FUNCTION_BLOCK TcoObjectTest EXTENDS TcoCore.TcoObject
VAR
	_myIdentity				:	ULINT;
	_myContextIdentity		:	ULINT;
	_myContextStartCount 	:	ULINT;
	_myContextEndCount		:	ULINT;
	_myParentIdentity		:	ULINT;
	_tcoTaskTest_A			:	TcoTaskTest(THIS^);
	_tcoTaskTest_B			:	TcoTaskTest(THIS^);
	_tcoStateTest_A			:	TcoStateTest(THIS^, eRestoreMode.AutoRestoreMembers);
	_tcoStateTest_B			:	TcoStateTest(THIS^, eRestoreMode.None);
	// Object equality
	_tcoObjectEqualsTestObj1 	:   TcoObjectEqualsTest(THIS^);
	_tcoObjectEqualsTestObj2 	:   TcoObjectEqualsTest(THIS^);
END_VAR

{attribute 'TcRpcEnable'}
METHOD INTERNAL CallTaskInstancies
_tcoTaskTest_A();

_tcoTaskTest_B();
END_METHOD

{attribute 'TcRpcEnable'}
METHOD PUBLIC EqualsOverrideTest : BOOL
EqualsOverrideTest := _tcoObjectEqualsTestObj1.EqualsTo(_tcoObjectEqualsTestObj2);
END_METHOD

{attribute 'TcRpcEnable'}
METHOD PUBLIC EqualsTest : BOOL
VAR_INPUT
    _case : INT;
END_VAR

VAR
    referenceTo_a_TcoStateTest : REFERENCE TO TcoStateTest;
END_VAR
CASE _case OF
    0:
        referenceTo_a_TcoStateTest REF= _tcoStateTest_A;
        EqualsTest := _tcoStateTest_A.EqualsTo(referenceTo_a_TcoStateTest);
    1:
        EqualsTest := _tcoStateTest_A.EqualsTo(_tcoStateTest_B);
    4:
        EqualsTest := _tcoStateTest_B.EqualsTo(_tcoStateTest_A);
    2:
        EqualsTest := _tcoObjectEqualsTestObj1.EqualsTo(_tcoObjectEqualsTestObj1);
    3:
        EqualsTest := _tcoObjectEqualsTestObj1.EqualsTo(_tcoObjectEqualsTestObj2);
END_CASE
END_METHOD

{attribute 'TcRpcEnable'}
METHOD INTERNAL ReadOutIdentities
_myIdentity			:=	THIS^.Identity;

_myContextIdentity	:=	THIS^.Context.Identity;
		
_myContextStartCount :=	THIS^.Context.StartCycleCount;

_myContextEndCount	:=	THIS^.Context.EndCycleCount;

_myParentIdentity	:=	THIS^.Parent.Identity;
END_METHOD

END_FUNCTION_BLOCK

(* stored: Version 1.1.0.1
   POU TcoObjectTest: Id {e84228ff-9c33-47a4-a38e-640688a82a88}, SpecialFunc None
   Method CallTaskInstancies: Id {ca9ba4d2-6103-4337-95bc-465f8f83317e}
   Method EqualsOverrideTest: Id {ee60d2fd-b5db-0d20-0c27-57a751cde2ce}
   Method EqualsTest: Id {9f06ff61-1678-0fe4-0121-54cfb8b16218}
   Method ReadOutIdentities: Id {b42bfa48-43e7-40ad-83bf-1125b1638f9d} *)
